(* IEC 61131-3 sources: beebread/doc/isa88, 7 files *)

(* ---- isa88_phase.st ---- *)
(*
 * ISA-88 phase template: the lowest procedural element, the one that runs
 * equipment. ISA88_PHASE wraps ISA88_STATE_MACHINE and adds what a phase's
 * equipment logic needs from it. A phase is written by composition:
 *
 *   FUNCTION_BLOCK PH_HEAT
 *     VAR ph : ISA88_PHASE; END_VAR
 *     ph(Start := cmdStart, Hold := cmdHold, FailCode := fault);
 *     CASE ph.State OF
 *       ISA88_RUNNING:
 *         IF ph.Entry THEN heater := TRUE; END_IF;
 *         IF temp >= setpoint THEN ph.Done(); END_IF;
 *       ISA88_HOLDING:
 *         heater := FALSE;
 *         ph.Done();
 *     END_CASE
 *
 * Each scan the phase logic calls ph first, then runs the logic of ph.State.
 *   Done()    : called by the logic when the current Running or transient
 *               state's work is finished (SC). The next call of ph takes it
 *               and forgets it, so it never carries into the next state.
 *               A transient state whose logic never calls Done stays in it.
 *   Entry     : TRUE on the first scan the logic runs a state; use it to
 *               start that state's work (open a valve, latch a restart step).
 *   StateTime : time spent in the current state, for timeouts.
 *   FailCode  : non-zero while the equipment has a failure. It holds the
 *               phase (Running, Pausing, Paused and Restarting accept Hold),
 *               so a Restart while the failure is still there holds again.
 *               The first code is latched in Failure until the phase is
 *               back in Idle.
 *
 * Commands are pulses, as for ISA88_STATE_MACHINE.
 *
 * Modes (ISA-88 procedural modes) decide how the logic moves from one step
 * to the next. The logic asks with Advance(condition):
 *
 *   ISA88_RUNNING:
 *     IF ph.JumpRequest THEN step := ph.JumpTarget;
 *     ELSIF ph.Advance(temp >= setpoint) THEN step := step + 1;
 *     END_IF;
 *
 *   Mode        : ISA88_AUTOMATIC (the default), ISA88_SEMI_AUTOMATIC or
 *                 ISA88_MANUAL. It may change at any time; another value
 *                 is ignored and ActiveMode keeps the last valid one.
 *   Advance(c)  : TRUE when the logic may take its next step.
 *                   Automatic      : when c is TRUE.
 *                   Semi-automatic : when c is TRUE and the operator
 *                                    presses Proceed.
 *                   Manual         : when the operator presses Proceed,
 *                                    whatever c is.
 *                 One Proceed allows one step.
 *   Waiting     : the logic is waiting on Proceed (Semi-automatic with its
 *                 condition met, or Manual).
 *   Jump        : Manual only: JumpRequest is TRUE for one scan, and the
 *                 logic moves to JumpTarget (JumpStep when Jump was pressed).
 *
 * Proceed and Jump act on their rising edge. Done() is not tied to a mode:
 * holding, stopping and aborting finish on their own in every mode, and a
 * step that should wait for the operator writes IF ph.Advance(c) THEN
 * ph.Done(); END_IF.
 *)
VAR_GLOBAL CONSTANT
	ISA88_IDLE       : INT := 1;
	ISA88_RUNNING    : INT := 2;
	ISA88_COMPLETE   : INT := 3;
	ISA88_PAUSING    : INT := 4;
	ISA88_PAUSED     : INT := 5;
	ISA88_HOLDING    : INT := 6;
	ISA88_HELD       : INT := 7;
	ISA88_RESTARTING : INT := 8;
	ISA88_STOPPING   : INT := 9;
	ISA88_STOPPED    : INT := 10;
	ISA88_ABORTING   : INT := 11;
	ISA88_ABORTED    : INT := 12;

	ISA88_AUTOMATIC      : INT := 1;
	ISA88_SEMI_AUTOMATIC : INT := 2;
	ISA88_MANUAL         : INT := 3;
END_VAR

FUNCTION_BLOCK ISA88_PHASE
	VAR_INPUT
		Start    : BOOL;
		Pause    : BOOL;
		Resume   : BOOL;
		Hold     : BOOL;
		Restart  : BOOL;
		Stop     : BOOL;
		Abort    : BOOL;
		Reset    : BOOL;
		FailCode : DINT; (* non-zero: equipment failure *)
		Mode     : INT := 1; (* ISA88_AUTOMATIC *)
		Proceed  : BOOL;
		Jump     : BOOL;
		JumpStep : INT;
	END_VAR
	VAR_OUTPUT
		State       : INT;
		Entry       : BOOL;
		StateTime   : TIME;
		Failure     : DINT;
		IsQuiescent : BOOL;
		IsTransient : BOOL;
		IsFinal     : BOOL;
		ActiveMode  : INT := 1; (* ISA88_AUTOMATIC *)
		Waiting     : BOOL;
		JumpRequest : BOOL;
		JumpTarget  : INT;
	END_VAR
	VAR
		sm          : ISA88_STATE_MACHINE;
		complete    : BOOL; (* Done was called since the last scan *)
		lastState   : INT;
		inState     : TON;
		proceedEdge : R_TRIG;
		jumpEdge    : R_TRIG;
		proceeding  : BOOL; (* a Proceed this scan not yet used by Advance *)
	END_VAR

	(* The current state's work is finished (SC). *)
	METHOD Done : BOOL
		complete := TRUE;
		Done := TRUE;
	END_METHOD

	(* May the logic take its next step, its condition being Cond? *)
	METHOD Advance : BOOL
		VAR_INPUT
			Cond : BOOL;
		END_VAR
		IF ActiveMode = ISA88_AUTOMATIC THEN
			Advance := Cond;
		ELSIF ActiveMode = ISA88_SEMI_AUTOMATIC AND NOT Cond THEN
			Advance := FALSE;
		ELSE
			Advance := proceeding;
			proceeding := FALSE;
			Waiting := NOT Advance;
		END_IF;
	END_METHOD

	sm(Start := Start, Pause := Pause, Resume := Resume,
	   Hold := Hold OR FailCode <> 0, Restart := Restart,
	   Stop := Stop, Abort := Abort, Reset := Reset, SC := complete);
	complete := FALSE;

	State := sm.State;
	IsQuiescent := sm.IsQuiescent;
	IsTransient := sm.IsTransient;
	IsFinal := sm.IsFinal;

	Entry := State <> lastState;
	lastState := State;
	inState(IN := NOT Entry, PT := T#24D);
	StateTime := inState.ET;

	IF State = ISA88_IDLE THEN
		Failure := 0;
	ELSIF FailCode <> 0 AND Failure = 0 THEN
		Failure := FailCode;
	END_IF;

	IF Mode = ISA88_AUTOMATIC OR Mode = ISA88_SEMI_AUTOMATIC OR Mode = ISA88_MANUAL THEN
		ActiveMode := Mode;
	END_IF;
	proceedEdge(CLK := Proceed);
	proceeding := proceedEdge.Q AND ActiveMode <> ISA88_AUTOMATIC;
	jumpEdge(CLK := Jump);
	JumpRequest := jumpEdge.Q AND ActiveMode = ISA88_MANUAL;
	IF JumpRequest THEN
		JumpTarget := JumpStep;
	END_IF;
	Waiting := FALSE; (* until Advance says otherwise this scan *)
END_FUNCTION_BLOCK

(* ---- isa88_phase_mode_test.st ---- *)
(* Unit tests for ISA88_PHASE modes:
   beedance -test isa88_state_machine.st isa88_phase.st isa88_phase_mode_test.st *)

(* A phase whose Running has steps 1 to 3. Each step's condition is Ready;
   after step 3 the phase is done. *)
FUNCTION_BLOCK PH_DEMO_STEPS
	VAR_INPUT
		Start    : BOOL;
		Reset    : BOOL;
		Mode     : INT := 1;
		Proceed  : BOOL;
		Jump     : BOOL;
		JumpStep : INT;
		Ready    : BOOL;
	END_VAR
	VAR_OUTPUT
		State      : INT;
		Step       : INT := 1;
		Waiting    : BOOL;
		ActiveMode : INT;
	END_VAR
	VAR
		ph : ISA88_PHASE;
	END_VAR
	ph(Start := Start, Reset := Reset, Mode := Mode, Proceed := Proceed, Jump := Jump, JumpStep := JumpStep);
	CASE ph.State OF
		ISA88_IDLE:
			IF ph.Entry THEN Step := 1; END_IF;
		ISA88_RUNNING:
			IF ph.JumpRequest THEN
				Step := ph.JumpTarget;
			ELSIF ph.Advance(Ready) THEN
				IF Step >= 3 THEN ph.Done(); ELSE Step := Step + 1; END_IF;
			END_IF;
	END_CASE
	State := ph.State;
	Waiting := ph.Waiting;
	ActiveMode := ph.ActiveMode;
END_FUNCTION_BLOCK

(* Automatic: a step is taken as soon as its condition is met; Proceed and
   Jump do nothing *)
PROGRAM TEST_MODE_Automatic
	VAR_OUTPUT
		failures : INT;
		message  : STRING;
		done     : BOOL;
	END_VAR
	VAR
		p    : PH_DEMO_STEPS;
		step : INT;
		ok   : BOOL;
	END_VAR
	ok := TRUE;
	CASE step OF
		0: p(); ok := p.State = ISA88_IDLE AND p.ActiveMode = ISA88_AUTOMATIC;
		1: p(Start := TRUE); ok := p.State = ISA88_RUNNING AND p.Step = 1 AND NOT p.Waiting;
		2: p(Start := FALSE, Proceed := TRUE, Jump := TRUE, JumpStep := 3); ok := p.Step = 1;
		3: p(Proceed := FALSE, Jump := FALSE, Ready := TRUE); ok := p.Step = 2 AND NOT p.Waiting;
		4: p(); ok := p.Step = 3;
		5: p(); ok := p.State = ISA88_RUNNING; (* step 3 met: Done *)
		6: p(); ok := p.State = ISA88_COMPLETE;
		   done := TRUE;
	END_CASE
	IF NOT ok THEN
		failures := failures + 1;
		message := CONCAT('wrong state after step ', INT_TO_STRING(step));
	END_IF;
	step := step + 1;
END_PROGRAM

(* Semi-automatic: a step needs its condition and a Proceed; one Proceed is
   one step; a Proceed before the condition is met is not kept *)
PROGRAM TEST_MODE_SemiAutomatic
	VAR_OUTPUT
		failures : INT;
		message  : STRING;
		done     : BOOL;
	END_VAR
	VAR
		p    : PH_DEMO_STEPS;
		step : INT;
		ok   : BOOL;
	END_VAR
	ok := TRUE;
	CASE step OF
		0: p(Mode := ISA88_SEMI_AUTOMATIC, Start := TRUE); ok := p.State = ISA88_RUNNING AND p.ActiveMode = ISA88_SEMI_AUTOMATIC AND NOT p.Waiting;
		1: p(Start := FALSE, Ready := TRUE); ok := p.Step = 1 AND p.Waiting;
		2: p(Proceed := TRUE); ok := p.Step = 2 AND NOT p.Waiting;
		3: p(); ok := p.Step = 2 AND p.Waiting; (* Proceed still held: no edge *)
		4: p(Proceed := FALSE, Ready := FALSE); ok := p.Step = 2 AND NOT p.Waiting;
		5: p(Proceed := TRUE); ok := p.Step = 2; (* condition not met *)
		6: p(Proceed := FALSE, Ready := TRUE); ok := p.Step = 2 AND p.Waiting; (* that Proceed was not kept *)
		7: p(Proceed := TRUE); ok := p.Step = 3;
		8: p(Proceed := FALSE); ok := p.Step = 3 AND p.Waiting;
		9: p(Proceed := TRUE); ok := p.State = ISA88_RUNNING; (* Done *)
		10: p(Proceed := FALSE); ok := p.State = ISA88_COMPLETE;
		    done := TRUE;
	END_CASE
	IF NOT ok THEN
		failures := failures + 1;
		message := CONCAT('wrong state after step ', INT_TO_STRING(step));
	END_IF;
	step := step + 1;
END_PROGRAM

(* Manual: the operator steps whatever the condition and may jump; the mode
   may change while running; an unknown mode is ignored *)
PROGRAM TEST_MODE_Manual
	VAR_OUTPUT
		failures : INT;
		message  : STRING;
		done     : BOOL;
	END_VAR
	VAR
		p    : PH_DEMO_STEPS;
		step : INT;
		ok   : BOOL;
	END_VAR
	ok := TRUE;
	CASE step OF
		0: p(Mode := ISA88_MANUAL, Start := TRUE); ok := p.State = ISA88_RUNNING AND p.Step = 1 AND p.Waiting;
		1: p(Start := FALSE, Proceed := TRUE); ok := p.Step = 2; (* Ready is FALSE *)
		2: p(Proceed := FALSE, Jump := TRUE, JumpStep := 1); ok := p.Step = 1;
		3: p(Jump := FALSE, Mode := 7); ok := p.ActiveMode = ISA88_MANUAL AND p.Step = 1;
		4: p(Proceed := TRUE); ok := p.Step = 2;
		5: p(Proceed := FALSE, Mode := ISA88_AUTOMATIC, Ready := TRUE); ok := p.ActiveMode = ISA88_AUTOMATIC AND p.Step = 3 AND NOT p.Waiting;
		6: p(Jump := TRUE, JumpStep := 1); ok := p.State = ISA88_RUNNING; (* no jump in Automatic: Done *)
		7: p(Jump := FALSE); ok := p.State = ISA88_COMPLETE AND p.Step = 3;
		   done := TRUE;
	END_CASE
	IF NOT ok THEN
		failures := failures + 1;
		message := CONCAT('wrong state after step ', INT_TO_STRING(step));
	END_IF;
	step := step + 1;
END_PROGRAM

(* ---- isa88_phase_test.st ---- *)
(* Unit tests for ISA88_PHASE:
   beedance -test isa88_state_machine.st isa88_phase.st isa88_phase_test.st *)

(* A heating phase written with the template: Running heats one degree a
   scan up to 5, Restarting takes 30 ms, the other transient states finish
   at once. Temp is kept across Hold and Restart, as a restart point. *)
FUNCTION_BLOCK PH_DEMO_HEAT
	VAR_INPUT
		Start   : BOOL;
		Hold    : BOOL;
		Restart : BOOL;
		Stop    : BOOL;
		Reset   : BOOL;
		Fault   : DINT;
	END_VAR
	VAR_OUTPUT
		Heater  : BOOL;
		Temp    : INT;
		State   : INT;
		Entry   : BOOL;
		Failure : DINT;
	END_VAR
	VAR
		ph : ISA88_PHASE;
	END_VAR
	ph(Start := Start, Hold := Hold, Restart := Restart, Stop := Stop, Reset := Reset, FailCode := Fault);
	CASE ph.State OF
		ISA88_IDLE:
			IF ph.Entry THEN Temp := 0; END_IF;
		ISA88_RUNNING:
			Heater := TRUE;
			Temp := Temp + 1;
			IF Temp >= 5 THEN ph.Done(); END_IF;
		ISA88_COMPLETE:
			Heater := FALSE;
		ISA88_HOLDING, ISA88_STOPPING, ISA88_ABORTING:
			Heater := FALSE;
			ph.Done();
		ISA88_RESTARTING:
			IF ph.StateTime >= T#30ms THEN ph.Done(); END_IF;
	END_CASE
	State := ph.State;
	Entry := ph.Entry;
	Failure := ph.Failure;
END_FUNCTION_BLOCK

(* Idle -> Running until the logic is done -> Complete -> Idle *)
PROGRAM TEST_PHASE_Complete
	VAR_OUTPUT
		failures : INT;
		message  : STRING;
		done     : BOOL;
	END_VAR
	VAR
		h    : PH_DEMO_HEAT;
		step : INT;
		ok   : BOOL;
	END_VAR
	ok := TRUE;
	CASE step OF
		0: h(); ok := h.State = ISA88_IDLE AND h.Entry;
		1: h(Start := TRUE); ok := h.State = ISA88_RUNNING AND h.Entry AND h.Heater AND h.Temp = 1;
		2: h(Start := FALSE); ok := h.State = ISA88_RUNNING AND NOT h.Entry AND h.Temp = 2;
		3: h(); ok := h.Temp = 3;
		4: h(); ok := h.Temp = 4;
		5: h(); ok := h.State = ISA88_RUNNING AND h.Temp = 5; (* logic sets Done *)
		6: h(); ok := h.State = ISA88_COMPLETE AND h.Entry AND NOT h.Heater;
		7: h(); ok := h.State = ISA88_COMPLETE AND NOT h.Entry;
		8: h(Reset := TRUE); ok := h.State = ISA88_IDLE AND h.Temp = 0;
		   done := TRUE;
	END_CASE
	IF NOT ok THEN
		failures := failures + 1;
		message := CONCAT('wrong state after step ', INT_TO_STRING(step));
	END_IF;
	step := step + 1;
END_PROGRAM

(* Done does not carry into the next state; Restarting waits on StateTime;
   Running resumes where it was held *)
PROGRAM TEST_PHASE_HoldRestart
	VAR_OUTPUT
		failures : INT;
		message  : STRING;
		done     : BOOL;
	END_VAR
	VAR
		h     : PH_DEMO_HEAT;
		step  : INT;
		ok    : BOOL;
		next  : BOOL;
		waits : INT;
	END_VAR
	ok := TRUE;
	next := TRUE;
	CASE step OF
		0: h(Start := TRUE); ok := h.State = ISA88_RUNNING AND h.Temp = 1;
		1: h(Start := FALSE, Hold := TRUE); ok := h.State = ISA88_HOLDING AND NOT h.Heater;
		2: h(Hold := FALSE); ok := h.State = ISA88_HELD;
		3: h(); ok := h.State = ISA88_HELD; (* Holding's Done was cleared *)
		4: h(Restart := TRUE); ok := h.State = ISA88_RESTARTING;
		5: h(Restart := FALSE); ok := h.State = ISA88_RESTARTING;
		6: h(); ok := h.State = ISA88_RESTARTING;
		7: h();
		   IF h.State = ISA88_RESTARTING THEN
		       waits := waits + 1;
		       ok := waits < 10;
		       next := FALSE;
		   ELSE
		       ok := h.State = ISA88_RUNNING AND h.Temp = 2;
		       done := TRUE;
		   END_IF;
	END_CASE
	IF NOT ok THEN
		failures := failures + 1;
		message := CONCAT('wrong state after step ', INT_TO_STRING(step));
		done := TRUE;
	END_IF;
	IF next THEN step := step + 1; END_IF;
END_PROGRAM

(* A failure holds the phase, Restart holds again while it lasts, Failure
   keeps the first code until Idle *)
PROGRAM TEST_PHASE_Failure
	VAR_OUTPUT
		failures : INT;
		message  : STRING;
		done     : BOOL;
	END_VAR
	VAR
		h    : PH_DEMO_HEAT;
		step : INT;
		ok   : BOOL;
	END_VAR
	ok := TRUE;
	CASE step OF
		0: h(Start := TRUE); ok := h.State = ISA88_RUNNING AND h.Failure = 0;
		1: h(Start := FALSE, Fault := 42); ok := h.State = ISA88_HOLDING AND h.Failure = 42;
		2: h(Fault := 99); ok := h.State = ISA88_HELD AND h.Failure = 42;
		3: h(Restart := TRUE); ok := h.State = ISA88_RESTARTING;
		4: h(Restart := FALSE); ok := h.State = ISA88_HOLDING; (* failure still there *)
		5: h(Fault := 0); ok := h.State = ISA88_HELD AND h.Failure = 42;
		6: h(Restart := TRUE); ok := h.State = ISA88_RESTARTING;
		7: h(Restart := FALSE, Stop := TRUE); ok := h.State = ISA88_STOPPING;
		8: h(Stop := FALSE); ok := h.State = ISA88_STOPPED AND h.Failure = 42;
		9: h(Reset := TRUE); ok := h.State = ISA88_IDLE AND h.Failure = 0;
		   done := TRUE;
	END_CASE
	IF NOT ok THEN
		failures := failures + 1;
		message := CONCAT('wrong state after step ', INT_TO_STRING(step));
	END_IF;
	step := step + 1;
END_PROGRAM

(* ---- isa88_sequencer.st ---- *)
(*
 * ISA-88 sequencer: up to 32 steps (0 to 31) run one after the other,
 * forward (0, 1, 2 ...) or in reverse (Count-1 ... 1, 0). Each step is an
 * ISA-88 phase (ISA88_PHASE, so an ISA88_STATE_MACHINE) with three times:
 *
 *   Starting : StartTime after the step starts
 *   Running  : then RunTime
 *   Stopping : then StopTime; the step is then Complete and the next one
 *              starts.
 *
 *   seq(Forward := pbFwd, Hold := pbHold, Count := 3,
 *       StartTime := tStart, RunTime := tRun, StopTime := tStop);
 *   motor1 := seq.Running[0];
 *
 * Commands are pulses, as for ISA88_STATE_MACHINE.
 *   Forward, Reverse : in Idle, start the sequence in that direction.
 *                      While it runs, change the direction: the running
 *                      step finishes and the next one is picked in the new
 *                      direction (Reverse from step 0, or Forward from the
 *                      last step, then completes the sequence).
 *   Pause, Resume, Hold, Restart, Stop, Abort
 *                    : go to the running step and act as ISA-88 says. A
 *                      command given between two steps waits for the next
 *                      one; Stop or Abort there ends the sequence at once.
 *   Reset            : from Complete, Stopped or Aborted back to Idle.
 *   Count            : steps in use, 0 to 32; it may change while the
 *                      sequence runs. 0 steps complete at once.
 *
 * State is the ISA-88 state of the sequence: Idle, then the running step's
 * state, then Complete, Stopped or Aborted. A Stop runs what is left of the
 * step's StopTime (all of it if the step had not reached Stopping); Pausing,
 * Holding, Restarting and Aborting finish at once. Held or Paused, a step's
 * time stands still, and Restart or Resume carry on from where it was.
 *
 * The order of the steps is a Sequential Function Chart, SEQ_CHART. Each
 * scan ISA88_SEQUENCER calls every step once, as the chart asked, then the
 * chart, on the steps' states. (A chart action that called the steps would
 * run them twice in a scan in which the chart moves.) A step starts the
 * scan after the chart picks it.
 *)

(* One step: an ISA-88 phase whose Running is Starting, Running and
   Stopping, timed. *)
FUNCTION_BLOCK SEQ_STEP
	VAR_INPUT
		Start     : BOOL;
		Pause     : BOOL;
		Resume    : BOOL;
		Hold      : BOOL;
		Restart   : BOOL;
		Stop      : BOOL;
		Abort     : BOOL;
		Reset     : BOOL;
		StartTime : TIME;
		RunTime   : TIME;
		StopTime  : TIME;
	END_VAR
	VAR_OUTPUT
		State    : INT;
		Starting : BOOL;
		Running  : BOOL;
		Stopping : BOOL;
		Elapsed  : TIME; (* time run in Starting, Running and Stopping *)
	END_VAR
	VAR
		ph       : ISA88_PHASE;
		base     : TIME; (* Elapsed when Running was entered *)
		stopLeft : TIME; (* what a Stop has left to run *)
	END_VAR
	ph(Start := Start, Pause := Pause, Resume := Resume, Hold := Hold,
	   Restart := Restart, Stop := Stop, Abort := Abort, Reset := Reset);
	Starting := FALSE;
	Running := FALSE;
	Stopping := FALSE;
	CASE ph.State OF
		ISA88_IDLE:
			Elapsed := T#0s;
		ISA88_RUNNING:
			IF ph.Entry THEN base := Elapsed; END_IF;
			Elapsed := base + ph.StateTime;
			IF Elapsed < StartTime THEN
				Starting := TRUE;
			ELSIF Elapsed < StartTime + RunTime THEN
				Running := TRUE;
			ELSIF Elapsed < StartTime + RunTime + StopTime THEN
				Stopping := TRUE;
			ELSE
				ph.Done();
			END_IF;
		ISA88_STOPPING:
			IF ph.Entry THEN
				IF Elapsed >= StartTime + RunTime + StopTime THEN
					stopLeft := T#0s;
				ELSIF Elapsed > StartTime + RunTime THEN
					stopLeft := StartTime + RunTime + StopTime - Elapsed;
				ELSE
					stopLeft := StopTime;
				END_IF;
			END_IF;
			IF ph.StateTime >= stopLeft THEN
				ph.Done();
			ELSE
				Stopping := TRUE;
			END_IF;
		ISA88_PAUSING, ISA88_HOLDING, ISA88_RESTARTING, ISA88_ABORTING:
			ph.Done();
	END_CASE
	State := ph.State;
END_FUNCTION_BLOCK

(* The order of the steps. StepState is the state of step Index; the
   chart asks for StepStart and StepReset on step Index. StopReq and
   AbortReq are a Stop or Abort no step has taken yet. *)
FUNCTION_BLOCK SEQ_CHART
	VAR_INPUT
		Go        : BOOL; (* Forward or Reverse *)
		Reversing : BOOL;
		Count     : INT;
		StepState : INT;
		StopReq   : BOOL;
		AbortReq  : BOOL;
		Reset     : BOOL;
	END_VAR
	VAR_OUTPUT
		Index     : INT := -1; (* the step in use; -1: none *)
		StepStart : BOOL;
		StepReset : BOOL;
		Busy      : BOOL; (* from the first step's start to the last step's end *)
		State     : INT := 1; (* ISA88_IDLE; while Busy, see the step *)
	END_VAR
	VAR
		NextIndex : INT;
		HasNext   : BOOL;
	END_VAR

	ACTION A_Idle:
		State := ISA88_IDLE;
		Index := -1;
		IF Reversing THEN NextIndex := Count - 1; ELSE NextIndex := 0; END_IF;
	END_ACTION
	ACTION A_Enter:
		Index := NextIndex;
		State := ISA88_RUNNING;
	END_ACTION
	ACTION A_Look:
		IF Reversing THEN
			NextIndex := MIN(Index, Count) - 1;
		ELSE
			NextIndex := Index + 1;
		END_IF;
		HasNext := NextIndex >= 0 AND NextIndex < Count;
	END_ACTION
	ACTION A_Complete:
		State := ISA88_COMPLETE;
		Index := -1;
	END_ACTION
	ACTION A_Stopped:
		State := ISA88_STOPPED;
	END_ACTION
	ACTION A_Aborted:
		State := ISA88_ABORTED;
	END_ACTION

	INITIAL_STEP S_Idle: A_Idle(N); END_STEP
	TRANSITION FROM S_Idle TO S_Start := Go AND Count > 0; END_TRANSITION
	TRANSITION FROM S_Idle TO S_Complete := Go AND Count <= 0; END_TRANSITION

	(* Start step Index; it has started once it leaves Idle. *)
	STEP S_Start: A_Enter(P); StepStart(N); Busy(N); END_STEP
	TRANSITION FROM S_Start TO S_Run := StepState <> ISA88_IDLE; END_TRANSITION

	(* The step runs, through whatever commands it is given, to an end. *)
	STEP S_Run: Busy(N); END_STEP
	TRANSITION FROM S_Run TO S_Next := StepState = ISA88_COMPLETE; END_TRANSITION
	TRANSITION FROM S_Run TO S_Stopped := StepState = ISA88_STOPPED; END_TRANSITION
	TRANSITION FROM S_Run TO S_Aborted := StepState = ISA88_ABORTED; END_TRANSITION

	(* Reset the finished step, then start the next one, if there is one. *)
	STEP S_Next: StepReset(N); A_Look(N); Busy(N); END_STEP
	TRANSITION FROM S_Next TO S_Aborted := AbortReq; END_TRANSITION
	TRANSITION FROM S_Next TO S_Stopped := StopReq AND NOT AbortReq; END_TRANSITION
	TRANSITION FROM S_Next TO S_Start := StepState = ISA88_IDLE AND HasNext AND NOT StopReq AND NOT AbortReq; END_TRANSITION
	TRANSITION FROM S_Next TO S_Complete := StepState = ISA88_IDLE AND NOT HasNext AND NOT StopReq AND NOT AbortReq; END_TRANSITION

	STEP S_Complete: A_Complete(N); END_STEP
	TRANSITION FROM S_Complete TO S_Idle := Reset; END_TRANSITION

	STEP S_Stopped: A_Stopped(N); END_STEP
	TRANSITION FROM S_Stopped TO S_Idle := Reset; END_TRANSITION

	STEP S_Aborted: A_Aborted(N); END_STEP
	TRANSITION FROM S_Aborted TO S_Idle := Reset; END_TRANSITION
END_FUNCTION_BLOCK

FUNCTION_BLOCK ISA88_SEQUENCER
	VAR_INPUT
		Forward   : BOOL;
		Reverse   : BOOL;
		Pause     : BOOL;
		Resume    : BOOL;
		Hold      : BOOL;
		Restart   : BOOL;
		Stop      : BOOL;
		Abort     : BOOL;
		Reset     : BOOL;
		Count     : INT; (* steps in use, 0 to 32 *)
		StartTime : ARRAY[0..31] OF TIME;
		RunTime   : ARRAY[0..31] OF TIME;
		StopTime  : ARRAY[0..31] OF TIME;
	END_VAR
	VAR_OUTPUT
		State     : INT := 1; (* ISA88_IDLE *)
		Index     : INT := -1; (* the step in use; -1: none *)
		Reversing : BOOL;
		Busy      : BOOL;
		Starting  : ARRAY[0..31] OF BOOL;
		Running   : ARRAY[0..31] OF BOOL;
		Stopping  : ARRAY[0..31] OF BOOL;
		StepState : ARRAY[0..31] OF INT;
	END_VAR
	VAR
		chart    : SEQ_CHART;
		steps    : ARRAY[0..31] OF SEQ_STEP;
		n        : INT;
		i        : INT;
		resetAll : BOOL;
		was      : INT; (* the state of step Index before this scan's call *)
		taken    : BOOL; (* step Index can take the pending commands *)
		pauseReq : BOOL;
		holdReq  : BOOL;
		stopReq  : BOOL;
		abortReq : BOOL;
	END_VAR
	n := LIMIT(0, Count, 32);
	IF Forward THEN
		Reversing := FALSE;
	ELSIF Reverse THEN
		Reversing := TRUE;
	END_IF;

	(* Commands wait while no step can take them: between two steps the
	   finished one is Complete and the next one Idle. *)
	IF chart.Busy THEN
		pauseReq := (pauseReq OR Pause) AND NOT Resume;
		holdReq := (holdReq OR Hold) AND NOT Restart;
		stopReq := stopReq OR Stop;
		abortReq := abortReq OR Abort;
	ELSE
		pauseReq := FALSE;
		holdReq := FALSE;
		stopReq := FALSE;
		abortReq := FALSE;
	END_IF;
	resetAll := Reset AND NOT chart.Busy;

	(* The steps first, as the chart asked last scan, then the chart, on
	   the steps as they are now. *)
	Index := chart.Index;
	Busy := chart.Busy;
	IF Index >= 0 AND Index <= 31 THEN
		was := steps[Index].State;
	ELSE
		was := ISA88_IDLE;
	END_IF;
	taken := was <> ISA88_IDLE AND was <> ISA88_COMPLETE;
	FOR i := 0 TO 31 DO
		IF i = Index AND Busy THEN
			steps[i](Start := chart.StepStart, Pause := pauseReq, Resume := Resume,
			         Hold := holdReq, Restart := Restart, Stop := stopReq,
			         Abort := abortReq, Reset := chart.StepReset OR resetAll,
			         StartTime := StartTime[i], RunTime := RunTime[i], StopTime := StopTime[i]);
		ELSE
			steps[i](Start := FALSE, Pause := FALSE, Resume := FALSE, Hold := FALSE,
			         Restart := FALSE, Stop := FALSE, Abort := FALSE, Reset := resetAll,
			         StartTime := StartTime[i], RunTime := RunTime[i], StopTime := StopTime[i]);
		END_IF;
		Starting[i] := steps[i].Starting;
		Running[i] := steps[i].Running;
		Stopping[i] := steps[i].Stopping;
		StepState[i] := steps[i].State;
	END_FOR;
	IF taken THEN
		pauseReq := FALSE;
		holdReq := FALSE;
	END_IF;

	IF Index >= 0 AND Index <= 31 THEN
		was := steps[Index].State;
	ELSE
		was := ISA88_IDLE;
	END_IF;
	chart(Go := Forward OR Reverse, Reversing := Reversing, Count := n,
	      StepState := was, StopReq := stopReq, AbortReq := abortReq,
	      Reset := Reset);
	Index := chart.Index;
	Busy := chart.Busy;

	IF Busy AND Index >= 0 AND Index <= 31 THEN
		State := steps[Index].State;
		IF State = ISA88_IDLE OR State = ISA88_COMPLETE THEN
			State := ISA88_RUNNING; (* between two steps *)
		END_IF;
	ELSE
		State := chart.State;
	END_IF;
END_FUNCTION_BLOCK

(* ---- isa88_sequencer_test.st ---- *)
(* Unit tests for ISA88_SEQUENCER:
   beedance -test isa88_state_machine.st isa88_phase.st isa88_sequencer.st isa88_sequencer_test.st

   The test runner scans every 10 ms of simulated time. *)

(* Records the order the steps run in. *)
FUNCTION_BLOCK SEQ_TRACE
	VAR_INPUT
		Index : INT;
	END_VAR
	VAR_OUTPUT
		Order     : ARRAY[0..39] OF INT;
		Runs      : INT;
		Ascending : BOOL; (* ran 0, 1, 2 ... *)
	END_VAR
	VAR
		last : INT := -1;
		k    : INT;
	END_VAR
	IF Index <> last AND Index >= 0 AND Runs <= 39 THEN
		Order[Runs] := Index;
		Runs := Runs + 1;
	END_IF;
	last := Index;
	Ascending := TRUE;
	FOR k := 0 TO Runs - 1 DO
		IF Order[k] <> k THEN Ascending := FALSE; END_IF;
	END_FOR;
END_FUNCTION_BLOCK

(* Sets the same times on the first n steps. *)
FUNCTION_BLOCK SEQ_TIMES
	VAR_INPUT
		n     : INT;
		start : TIME;
		run   : TIME;
		stop  : TIME;
	END_VAR
	VAR_OUTPUT
		StartTime : ARRAY[0..31] OF TIME;
		RunTime   : ARRAY[0..31] OF TIME;
		StopTime  : ARRAY[0..31] OF TIME;
	END_VAR
	VAR
		k : INT;
	END_VAR
	FOR k := 0 TO n - 1 DO
		StartTime[k] := start;
		RunTime[k] := run;
		StopTime[k] := stop;
	END_FOR;
END_FUNCTION_BLOCK

(* Three steps forward: 0, 1, 2, each Starting, Running then Stopping,
   then Complete, then Reset to Idle *)
PROGRAM TEST_SEQ_Forward
	VAR_OUTPUT
		failures : INT;
		message  : STRING;
		done     : BOOL;
	END_VAR
	VAR
		seq      : ISA88_SEQUENCER;
		tm       : SEQ_TIMES;
		tr       : SEQ_TRACE;
		scan     : INT;
		sawStart : BOOL;
		sawRun   : BOOL;
		sawStop  : BOOL;
		overlap  : BOOL;
		on       : INT;
	END_VAR
	tm(n := 3, start := T#20ms, run := T#30ms, stop := T#20ms);
	seq(Forward := scan = 0, Reset := FALSE, Count := 3,
	    StartTime := tm.StartTime, RunTime := tm.RunTime, StopTime := tm.StopTime);
	tr(Index := seq.Index);
	IF seq.Starting[0] THEN sawStart := TRUE; END_IF;
	IF seq.Running[0] THEN sawRun := TRUE; END_IF;
	IF seq.Stopping[0] THEN sawStop := TRUE; END_IF;
	on := 0;
	IF seq.Starting[0] OR seq.Running[0] OR seq.Stopping[0] THEN on := on + 1; END_IF;
	IF seq.Starting[1] OR seq.Running[1] OR seq.Stopping[1] THEN on := on + 1; END_IF;
	IF seq.Starting[2] OR seq.Running[2] OR seq.Stopping[2] THEN on := on + 1; END_IF;
	IF on > 1 THEN overlap := TRUE; END_IF;
	IF scan = 0 AND NOT (seq.Busy AND seq.Index = 0 AND seq.State = ISA88_RUNNING) THEN
		failures := failures + 1; message := 'Forward did not start step 0'; done := TRUE;
	END_IF;
	IF seq.State = ISA88_COMPLETE AND NOT done THEN
		IF tr.Runs <> 3 OR tr.Order[0] <> 0 OR tr.Order[1] <> 1 OR tr.Order[2] <> 2 THEN
			failures := failures + 1; message := 'steps not run 0, 1, 2';
		ELSIF NOT (sawStart AND sawRun AND sawStop) THEN
			failures := failures + 1; message := 'step 0 missed a phase';
		ELSIF overlap THEN
			failures := failures + 1; message := 'two steps on at once';
		ELSIF seq.Busy OR seq.Index <> -1 THEN
			failures := failures + 1; message := 'Complete but busy';
		ELSE
			seq(Reset := TRUE);
			IF seq.State <> ISA88_IDLE OR seq.StepState[2] <> ISA88_IDLE THEN
				failures := failures + 1; message := 'Reset did not go to Idle';
			END_IF;
		END_IF;
		done := TRUE;
	END_IF;
	scan := scan + 1;
	IF scan > 200 AND NOT done THEN
		failures := failures + 1; message := 'never completed'; done := TRUE;
	END_IF;
END_PROGRAM

(* Step 0's phases follow its three times: 2 scans Starting, 3 Running,
   2 Stopping *)
PROGRAM TEST_SEQ_StepTimes
	VAR_OUTPUT
		failures : INT;
		message  : STRING;
		done     : BOOL;
	END_VAR
	VAR
		seq    : ISA88_SEQUENCER;
		scan   : INT;
		nStart : INT;
		nRun   : INT;
		nStop  : INT;
	END_VAR
	seq.StartTime[0] := T#20ms;
	seq.RunTime[0] := T#30ms;
	seq.StopTime[0] := T#20ms;
	seq(Forward := scan = 0, Count := 1);
	IF seq.Starting[0] THEN nStart := nStart + 1; END_IF;
	IF seq.Running[0] THEN nRun := nRun + 1; END_IF;
	IF seq.Stopping[0] THEN nStop := nStop + 1; END_IF;
	IF seq.State = ISA88_COMPLETE THEN
		IF nStart < 2 OR nStart > 3 OR nRun <> 3 OR nStop <> 2 THEN
			failures := failures + 1;
			message := CONCAT(CONCAT(CONCAT('scans Starting/Running/Stopping: ', INT_TO_STRING(nStart)),
			           CONCAT('/', INT_TO_STRING(nRun))), CONCAT('/', INT_TO_STRING(nStop)));
		END_IF;
		done := TRUE;
	END_IF;
	scan := scan + 1;
	IF scan > 100 AND NOT done THEN
		failures := failures + 1; message := 'never completed'; done := TRUE;
	END_IF;
END_PROGRAM

(* Reverse runs 2, 1, 0 *)
PROGRAM TEST_SEQ_Reverse
	VAR_OUTPUT
		failures : INT;
		message  : STRING;
		done     : BOOL;
	END_VAR
	VAR
		seq  : ISA88_SEQUENCER;
		tr   : SEQ_TRACE;
		scan : INT;
	END_VAR
	seq(Reverse := scan = 0, Count := 3);
	tr(Index := seq.Index);
	IF seq.State = ISA88_COMPLETE THEN
		IF NOT seq.Reversing OR tr.Runs <> 3 OR tr.Order[0] <> 2 OR tr.Order[1] <> 1 OR tr.Order[2] <> 0 THEN
			failures := failures + 1; message := 'steps not run 2, 1, 0';
		END_IF;
		done := TRUE;
	END_IF;
	scan := scan + 1;
	IF scan > 200 AND NOT done THEN
		failures := failures + 1; message := 'never completed'; done := TRUE;
	END_IF;
END_PROGRAM

(* Reverse while step 2 of 5 runs: 0, 1, 2, then back 1, 0 *)
PROGRAM TEST_SEQ_ChangeDirection
	VAR_OUTPUT
		failures : INT;
		message  : STRING;
		done     : BOOL;
	END_VAR
	VAR
		seq  : ISA88_SEQUENCER;
		tm   : SEQ_TIMES;
		tr   : SEQ_TRACE;
		scan : INT;
		sent : BOOL;
		rev  : BOOL;
	END_VAR
	tm(n := 5, run := T#30ms);
	rev := seq.Index = 2 AND NOT sent;
	IF rev THEN sent := TRUE; END_IF;
	seq(Forward := scan = 0, Reverse := rev, Count := 5, RunTime := tm.RunTime);
	tr(Index := seq.Index);
	IF seq.State = ISA88_COMPLETE THEN
		IF tr.Runs <> 5 OR tr.Order[0] <> 0 OR tr.Order[1] <> 1 OR tr.Order[2] <> 2
		   OR tr.Order[3] <> 1 OR tr.Order[4] <> 0 THEN
			failures := failures + 1; message := 'steps not run 0, 1, 2, 1, 0';
		END_IF;
		done := TRUE;
	END_IF;
	scan := scan + 1;
	IF scan > 300 AND NOT done THEN
		failures := failures + 1; message := 'never completed'; done := TRUE;
	END_IF;
END_PROGRAM

(* No steps: Complete at once; Reset back to Idle *)
PROGRAM TEST_SEQ_Empty
	VAR_OUTPUT
		failures : INT;
		message  : STRING;
		done     : BOOL;
	END_VAR
	VAR
		seq : ISA88_SEQUENCER;
		ok  : BOOL;
	END_VAR
	seq(Count := 0);
	ok := seq.State = ISA88_IDLE AND NOT seq.Busy;
	seq(Forward := TRUE);
	ok := ok AND seq.State = ISA88_COMPLETE AND seq.Index = -1 AND NOT seq.Busy;
	seq(Forward := FALSE, Reset := TRUE);
	ok := ok AND seq.State = ISA88_IDLE;
	IF NOT ok THEN
		failures := 1; message := 'empty sequence';
	END_IF;
	done := TRUE;
END_PROGRAM

(* All 32 steps, forward, with no times: each runs once, in order *)
PROGRAM TEST_SEQ_ThirtyTwo
	VAR_OUTPUT
		failures : INT;
		message  : STRING;
		done     : BOOL;
	END_VAR
	VAR
		seq  : ISA88_SEQUENCER;
		tr   : SEQ_TRACE;
		scan : INT;
	END_VAR
	seq(Forward := scan = 0, Count := 40); (* more than 32 is 32 *)
	tr(Index := seq.Index);
	IF seq.State = ISA88_COMPLETE THEN
		IF tr.Runs <> 32 OR NOT tr.Ascending THEN
			failures := failures + 1; message := 'steps not run 0 to 31';
		END_IF;
		done := TRUE;
	END_IF;
	scan := scan + 1;
	IF scan > 1000 AND NOT done THEN
		failures := failures + 1; message := 'never completed'; done := TRUE;
	END_IF;
END_PROGRAM

(* Hold while step 1 runs: Held, its time stands still; Restart carries on
   and the sequence completes *)
PROGRAM TEST_SEQ_HoldRestart
	VAR_OUTPUT
		failures : INT;
		message  : STRING;
		done     : BOOL;
	END_VAR
	VAR
		seq   : ISA88_SEQUENCER;
		tm    : SEQ_TIMES;
		tr    : SEQ_TRACE;
		scan  : INT;
		phase : INT;
		wait  : INT;
	END_VAR
	tm(n := 3, run := T#50ms);
	CASE phase OF
		0: seq(Forward := scan = 0, Count := 3, RunTime := tm.RunTime);
		   IF seq.Index = 1 AND seq.Running[1] THEN
		       seq(Hold := TRUE);
		       IF seq.State <> ISA88_HOLDING THEN
		           failures := failures + 1; message := 'Hold did not go to Holding'; done := TRUE;
		       END_IF;
		       phase := 1;
		   END_IF;
		1: seq(Hold := FALSE);
		   IF seq.State = ISA88_HELD THEN
		       wait := wait + 1;
		       IF seq.Running[1] OR seq.Index <> 1 THEN
		           failures := failures + 1; message := 'Held but running'; done := TRUE;
		       ELSIF wait = 10 THEN
		           seq(Restart := TRUE);
		           IF seq.State <> ISA88_RESTARTING THEN
		               failures := failures + 1; message := 'Restart did not go to Restarting'; done := TRUE;
		           END_IF;
		           phase := 2;
		       END_IF;
		   END_IF;
		2: seq(Restart := FALSE);
		   IF seq.State = ISA88_COMPLETE THEN
		       IF tr.Runs <> 3 THEN
		           failures := failures + 1; message := 'did not carry on to step 2';
		       END_IF;
		       done := TRUE;
		   END_IF;
	END_CASE
	tr(Index := seq.Index);
	scan := scan + 1;
	IF scan > 300 AND NOT done THEN
		failures := failures + 1; message := 'never completed'; done := TRUE;
	END_IF;
END_PROGRAM

(* Stop while step 0 runs: Stopping runs StopTime, then Stopped; step 1
   never starts; Reset makes every step Idle *)
PROGRAM TEST_SEQ_Stop
	VAR_OUTPUT
		failures : INT;
		message  : STRING;
		done     : BOOL;
	END_VAR
	VAR
		seq   : ISA88_SEQUENCER;
		scan  : INT;
		phase : INT;
		nStop : INT;
	END_VAR
	seq.RunTime[0] := T#100ms;
	seq.StopTime[0] := T#30ms;
	CASE phase OF
		0: seq(Forward := scan = 0, Count := 2);
		   IF scan = 3 THEN
		       seq(Stop := TRUE);
		       phase := 1;
		   END_IF;
		1: seq(Stop := FALSE);
		   IF seq.Stopping[0] THEN nStop := nStop + 1; END_IF;
		   IF seq.State = ISA88_STOPPED THEN
		       IF nStop <> 3 OR seq.StepState[1] <> ISA88_IDLE OR seq.Busy THEN
		           failures := failures + 1; message := CONCAT('wrong stop, scans Stopping: ', INT_TO_STRING(nStop));
		       END_IF;
		       seq(Reset := TRUE);
		       IF seq.State <> ISA88_IDLE OR seq.StepState[0] <> ISA88_IDLE THEN
		           failures := failures + 1; message := 'Reset did not go to Idle';
		       END_IF;
		       done := TRUE;
		   END_IF;
	END_CASE
	scan := scan + 1;
	IF scan > 100 AND NOT done THEN
		failures := failures + 1; message := 'never stopped'; done := TRUE;
	END_IF;
END_PROGRAM

(* Stop and Abort given between two steps are not lost *)
PROGRAM TEST_SEQ_BetweenSteps
	VAR_OUTPUT
		failures : INT;
		message  : STRING;
		done     : BOOL;
	END_VAR
	VAR
		a, b  : ISA88_SEQUENCER;
		scan  : INT;
		gapA  : BOOL;
		gapB  : BOOL;
		sentA : BOOL;
		sentB : BOOL;
	END_VAR
	(* the scan step 0 reports Complete, the chart is between steps *)
	gapA := a.StepState[0] = ISA88_COMPLETE AND NOT sentA;
	IF gapA THEN sentA := TRUE; END_IF;
	gapB := b.StepState[0] = ISA88_COMPLETE AND NOT sentB;
	IF gapB THEN sentB := TRUE; END_IF;
	a(Forward := scan = 0, Stop := gapA, Count := 3);
	b(Forward := scan = 0, Abort := gapB, Count := 3);
	IF scan = 40 THEN
		IF a.State <> ISA88_STOPPED OR a.StepState[1] = ISA88_RUNNING THEN
			failures := failures + 1; message := 'Stop between steps was lost';
		ELSIF b.State <> ISA88_ABORTED THEN
			failures := failures + 1; message := 'Abort between steps was lost';
		ELSIF NOT (sentA AND sentB) THEN
			failures := failures + 1; message := 'never between steps';
		END_IF;
		done := TRUE;
	END_IF;
	scan := scan + 1;
END_PROGRAM

(* Abort while a step runs: Aborted; Reset to Idle *)
PROGRAM TEST_SEQ_Abort
	VAR_OUTPUT
		failures : INT;
		message  : STRING;
		done     : BOOL;
	END_VAR
	VAR
		seq : ISA88_SEQUENCER;
		ok  : BOOL;
	END_VAR
	seq.RunTime[0] := T#1s;
	seq(Forward := TRUE, Count := 4);
	ok := seq.State = ISA88_RUNNING AND seq.Index = 0 AND NOT seq.Running[0]; (* starts next scan *)
	seq(Forward := FALSE);
	ok := ok AND seq.State = ISA88_RUNNING AND NOT seq.Starting[0] AND seq.Running[0];
	seq(Abort := TRUE);
	ok := ok AND seq.State = ISA88_ABORTING AND NOT seq.Running[0];
	seq(Abort := FALSE);
	ok := ok AND seq.State = ISA88_ABORTED;
	seq();
	ok := ok AND seq.State = ISA88_ABORTED AND NOT seq.Busy;
	seq(Reset := TRUE);
	ok := ok AND seq.State = ISA88_IDLE AND seq.StepState[0] = ISA88_IDLE;
	IF NOT ok THEN
		failures := 1; message := 'abort';
	END_IF;
	done := TRUE;
END_PROGRAM

(* ---- isa88_state_machine.st ---- *)
(*
 * ISA-88 (IEC 61512-1) procedural state machine as a Sequential Function Chart.
 *
 * One step per procedural state; one transition per arrow of the ISA-88
 * state diagram. Commands are inputs, pulsed by the caller for one scan.
 * SC (state complete) is raised by the procedural logic when the logic of
 * the current Running or transient state has finished.
 *
 *   Initial    : Idle
 *   Quiescent  : Idle, Paused, Held
 *   Transient  : Running, Pausing, Holding, Restarting, Stopping, Aborting
 *   Final      : Complete, Stopped, Aborted
 *
 * Which commands a state accepts (the nested boxes of the diagram):
 *   Pause  : Running
 *   Resume : Paused
 *   Hold   : Running, Pausing, Paused, Restarting
 *   Restart: Held
 *   Stop   : Running, Pausing, Paused, Holding, Held, Restarting
 *   Abort  : every state except Idle, Complete, Aborting and Aborted
 *   Reset  : Complete, Stopped, Aborted
 *
 * A step fires at most one transition per scan, so where a state accepts
 * more than one command they are ranked: Abort, Stop, Hold, Pause or
 * Resume or Restart, then SC.
 *
 * State codes (ISA-88 names no numbers; these are beebread's):
 *   1 Idle      2 Running   3 Complete
 *   4 Pausing   5 Paused    6 Holding   7 Held      8 Restarting
 *   9 Stopping 10 Stopped  11 Aborting 12 Aborted
 *)
FUNCTION_BLOCK ISA88_STATE_MACHINE
	VAR_INPUT
		Start   : BOOL;
		Pause   : BOOL;
		Resume  : BOOL;
		Hold    : BOOL;
		Restart : BOOL;
		Stop    : BOOL;
		Abort   : BOOL;
		Reset   : BOOL;
		SC      : BOOL; (* state complete *)
	END_VAR
	VAR_OUTPUT
		State       : INT;
		IsQuiescent : BOOL;
		IsTransient : BOOL;
		IsFinal     : BOOL;
	END_VAR

	ACTION A_Idle:
		State := 1; IsQuiescent := TRUE; IsTransient := FALSE; IsFinal := FALSE;
	END_ACTION
	ACTION A_Running:
		State := 2; IsQuiescent := FALSE; IsTransient := TRUE; IsFinal := FALSE;
	END_ACTION
	ACTION A_Complete:
		State := 3; IsQuiescent := FALSE; IsTransient := FALSE; IsFinal := TRUE;
	END_ACTION
	ACTION A_Pausing:
		State := 4; IsQuiescent := FALSE; IsTransient := TRUE; IsFinal := FALSE;
	END_ACTION
	ACTION A_Paused:
		State := 5; IsQuiescent := TRUE; IsTransient := FALSE; IsFinal := FALSE;
	END_ACTION
	ACTION A_Holding:
		State := 6; IsQuiescent := FALSE; IsTransient := TRUE; IsFinal := FALSE;
	END_ACTION
	ACTION A_Held:
		State := 7; IsQuiescent := TRUE; IsTransient := FALSE; IsFinal := FALSE;
	END_ACTION
	ACTION A_Restarting:
		State := 8; IsQuiescent := FALSE; IsTransient := TRUE; IsFinal := FALSE;
	END_ACTION
	ACTION A_Stopping:
		State := 9; IsQuiescent := FALSE; IsTransient := TRUE; IsFinal := FALSE;
	END_ACTION
	ACTION A_Stopped:
		State := 10; IsQuiescent := FALSE; IsTransient := FALSE; IsFinal := TRUE;
	END_ACTION
	ACTION A_Aborting:
		State := 11; IsQuiescent := FALSE; IsTransient := TRUE; IsFinal := FALSE;
	END_ACTION
	ACTION A_Aborted:
		State := 12; IsQuiescent := FALSE; IsTransient := FALSE; IsFinal := TRUE;
	END_ACTION

	(* ---- Initial state ---- *)
	INITIAL_STEP Idle: A_Idle(N); END_STEP
	TRANSITION FROM Idle TO Running := Start; END_TRANSITION

	(* ---- Running ---- *)
	STEP Running: A_Running(N); END_STEP
	TRANSITION FROM Running TO Aborting := Abort; END_TRANSITION
	TRANSITION FROM Running TO Stopping := Stop AND NOT Abort; END_TRANSITION
	TRANSITION FROM Running TO Holding := Hold AND NOT Stop AND NOT Abort; END_TRANSITION
	TRANSITION FROM Running TO Pausing := Pause AND NOT Hold AND NOT Stop AND NOT Abort; END_TRANSITION
	TRANSITION FROM Running TO Complete := SC AND NOT Pause AND NOT Hold AND NOT Stop AND NOT Abort; END_TRANSITION

	(* ---- Pause ---- *)
	STEP Pausing: A_Pausing(N); END_STEP
	TRANSITION FROM Pausing TO Aborting := Abort; END_TRANSITION
	TRANSITION FROM Pausing TO Stopping := Stop AND NOT Abort; END_TRANSITION
	TRANSITION FROM Pausing TO Holding := Hold AND NOT Stop AND NOT Abort; END_TRANSITION
	TRANSITION FROM Pausing TO Paused := SC AND NOT Hold AND NOT Stop AND NOT Abort; END_TRANSITION

	STEP Paused: A_Paused(N); END_STEP
	TRANSITION FROM Paused TO Aborting := Abort; END_TRANSITION
	TRANSITION FROM Paused TO Stopping := Stop AND NOT Abort; END_TRANSITION
	TRANSITION FROM Paused TO Holding := Hold AND NOT Stop AND NOT Abort; END_TRANSITION
	TRANSITION FROM Paused TO Running := Resume AND NOT Hold AND NOT Stop AND NOT Abort; END_TRANSITION

	(* ---- Hold ---- *)
	STEP Holding: A_Holding(N); END_STEP
	TRANSITION FROM Holding TO Aborting := Abort; END_TRANSITION
	TRANSITION FROM Holding TO Stopping := Stop AND NOT Abort; END_TRANSITION
	TRANSITION FROM Holding TO Held := SC AND NOT Stop AND NOT Abort; END_TRANSITION

	STEP Held: A_Held(N); END_STEP
	TRANSITION FROM Held TO Aborting := Abort; END_TRANSITION
	TRANSITION FROM Held TO Stopping := Stop AND NOT Abort; END_TRANSITION
	TRANSITION FROM Held TO Restarting := Restart AND NOT Stop AND NOT Abort; END_TRANSITION

	STEP Restarting: A_Restarting(N); END_STEP
	TRANSITION FROM Restarting TO Aborting := Abort; END_TRANSITION
	TRANSITION FROM Restarting TO Stopping := Stop AND NOT Abort; END_TRANSITION
	TRANSITION FROM Restarting TO Holding := Hold AND NOT Stop AND NOT Abort; END_TRANSITION
	TRANSITION FROM Restarting TO Running := SC AND NOT Hold AND NOT Stop AND NOT Abort; END_TRANSITION

	(* ---- Stop ---- *)
	STEP Stopping: A_Stopping(N); END_STEP
	TRANSITION FROM Stopping TO Aborting := Abort; END_TRANSITION
	TRANSITION FROM Stopping TO Stopped := SC AND NOT Abort; END_TRANSITION

	STEP Stopped: A_Stopped(N); END_STEP
	TRANSITION FROM Stopped TO Aborting := Abort; END_TRANSITION
	TRANSITION FROM Stopped TO Idle := Reset AND NOT Abort; END_TRANSITION

	(* ---- Abort ---- *)
	STEP Aborting: A_Aborting(N); END_STEP
	TRANSITION FROM Aborting TO Aborted := SC; END_TRANSITION

	STEP Aborted: A_Aborted(N); END_STEP
	TRANSITION FROM Aborted TO Idle := Reset; END_TRANSITION

	(* ---- Complete ---- *)
	STEP Complete: A_Complete(N); END_STEP
	TRANSITION FROM Complete TO Idle := Reset; END_TRANSITION
END_FUNCTION_BLOCK

(* ---- isa88_state_machine_test.st ---- *)
(* Unit tests for ISA88_STATE_MACHINE:
   beedance -test isa88_state_machine.st isa88_state_machine_test.st *)

(* Idle -> Running -> Complete -> Idle *)
PROGRAM TEST_ISA88_Complete
	VAR_OUTPUT
		failures : INT;
		message  : STRING;
		done     : BOOL;
	END_VAR
	VAR
		sm   : ISA88_STATE_MACHINE;
		step : INT;
		ok   : BOOL;
	END_VAR
	ok := TRUE;
	CASE step OF
		0: sm(); ok := ok AND sm.State = 1 AND sm.IsQuiescent;
		1: sm(Start := TRUE); ok := ok AND sm.State = 2 AND sm.IsTransient;
		2: sm(Start := FALSE); ok := ok AND sm.State = 2;
		3: sm(SC := TRUE); ok := ok AND sm.State = 3 AND sm.IsFinal;
		4: sm(SC := FALSE, Reset := TRUE); ok := ok AND sm.State = 1;
		5: sm(Reset := FALSE); ok := ok AND sm.State = 1;
		   done := TRUE;
	END_CASE
	IF NOT ok THEN
		failures := failures + 1;
		message := CONCAT('wrong state after step ', INT_TO_STRING(step));
	END_IF;
	step := step + 1;
END_PROGRAM

(* Running -> Pausing -> Paused -> Running -> Holding -> Held -> Restarting -> Running *)
PROGRAM TEST_ISA88_PauseHold
	VAR_OUTPUT
		failures : INT;
		message  : STRING;
		done     : BOOL;
	END_VAR
	VAR
		sm   : ISA88_STATE_MACHINE;
		step : INT;
		ok   : BOOL;
	END_VAR
	ok := TRUE;
	CASE step OF
		0: sm(Start := TRUE); ok := ok AND sm.State = 2;
		1: sm(Start := FALSE, Pause := TRUE); ok := ok AND sm.State = 4;
		2: sm(Pause := FALSE, SC := TRUE); ok := ok AND sm.State = 5 AND sm.IsQuiescent;
		3: sm(SC := FALSE, Resume := TRUE); ok := ok AND sm.State = 2;
		4: sm(Resume := FALSE, Hold := TRUE); ok := ok AND sm.State = 6;
		5: sm(Hold := FALSE, SC := TRUE); ok := ok AND sm.State = 7 AND sm.IsQuiescent;
		6: sm(SC := FALSE, Restart := TRUE); ok := ok AND sm.State = 8;
		7: sm(Restart := FALSE, Hold := TRUE); ok := ok AND sm.State = 6; (* Hold while Restarting *)
		8: sm(Hold := FALSE, SC := TRUE); ok := ok AND sm.State = 7;
		9: sm(SC := FALSE, Restart := TRUE); ok := ok AND sm.State = 8;
		10: sm(Restart := FALSE, SC := TRUE); ok := ok AND sm.State = 2;
		11: sm(SC := FALSE, Pause := TRUE); ok := ok AND sm.State = 4;
		12: sm(Pause := FALSE, Hold := TRUE); ok := ok AND sm.State = 6; (* Hold while Pausing *)
		    done := TRUE;
	END_CASE
	IF NOT ok THEN
		failures := failures + 1;
		message := CONCAT('wrong state after step ', INT_TO_STRING(step));
	END_IF;
	step := step + 1;
END_PROGRAM

(* Stop and Abort paths, command priority, and commands a state ignores *)
PROGRAM TEST_ISA88_StopAbort
	VAR_OUTPUT
		failures : INT;
		message  : STRING;
		done     : BOOL;
	END_VAR
	VAR
		sm   : ISA88_STATE_MACHINE;
		step : INT;
		ok   : BOOL;
	END_VAR
	ok := TRUE;
	CASE step OF
		0: sm(Stop := TRUE, Abort := TRUE, Hold := TRUE); ok := ok AND sm.State = 1; (* Idle ignores them *)
		1: sm(Stop := FALSE, Abort := FALSE, Hold := FALSE, Start := TRUE); ok := ok AND sm.State = 2;
		2: sm(Start := FALSE, Hold := TRUE, Stop := TRUE); ok := ok AND sm.State = 9; (* Stop beats Hold *)
		3: sm(Hold := FALSE, Stop := FALSE, SC := TRUE); ok := ok AND sm.State = 10 AND sm.IsFinal;
		4: sm(SC := FALSE, Abort := TRUE); ok := ok AND sm.State = 11; (* Abort from Stopped *)
		5: sm(Abort := FALSE, Reset := TRUE); ok := ok AND sm.State = 11; (* Aborting ignores Reset *)
		6: sm(Reset := FALSE, SC := TRUE); ok := ok AND sm.State = 12 AND sm.IsFinal;
		7: sm(SC := FALSE, Start := TRUE); ok := ok AND sm.State = 12; (* Aborted ignores Start *)
		8: sm(Start := FALSE, Reset := TRUE); ok := ok AND sm.State = 1;
		9: sm(Reset := FALSE, Start := TRUE); ok := ok AND sm.State = 2;
		10: sm(Start := FALSE, Stop := TRUE, Abort := TRUE); ok := ok AND sm.State = 11; (* Abort beats Stop *)
		11: sm(Stop := FALSE, Abort := FALSE, SC := TRUE); ok := ok AND sm.State = 12;
		12: sm(SC := FALSE, Reset := TRUE); ok := ok AND sm.State = 1;
		    done := TRUE;
	END_CASE
	IF NOT ok THEN
		failures := failures + 1;
		message := CONCAT('wrong state after step ', INT_TO_STRING(step));
	END_IF;
	step := step + 1;
END_PROGRAM
